(* IEC 61131-3 sources: ironplc/compiler/resources/test, 62 files *)

(* ---- first_steps_data_type_decl.st ---- *)
TYPE
  LOGLEVEL : (CRITICAL, WARNING, INFO, DEBUG) := INFO;
END_TYPE

(* ---- sized_string_contexts.st ---- *)
FUNCTION FUNC_WITH_VAR_STRING : INT
VAR_INPUT
    x : INT;
END_VAR
VAR
    buf : STRING[10];
    wbuf : WSTRING[20];
END_VAR
FUNC_WITH_VAR_STRING := 0;
END_FUNCTION

FUNCTION FUNC_WITH_VAR_CONSTANT_STRING : INT
VAR CONSTANT
    FILL : STRING[1] := '0';
    WFILL : WSTRING[1] := "0";
END_VAR
FUNC_WITH_VAR_CONSTANT_STRING := 0;
END_FUNCTION

FUNCTION FUNC_WITH_VAR_IN_OUT_STRING : INT
VAR_IN_OUT
    buf : STRING[255];
    wbuf : WSTRING[255];
END_VAR
FUNC_WITH_VAR_IN_OUT_STRING := 0;
END_FUNCTION

TYPE STRUCT_WITH_STRING :
STRUCT
    name : STRING[10];
    wname : WSTRING[20];
END_STRUCT;
END_TYPE

(* ---- strings.st ---- *)
TYPE
   TEXT_EXTENDED : STRING [1] := '�';
END_TYPE

(* ---- type_decl.st ---- *)
TYPE
   VALUES_ENUM : (VAL1, VAL2, VAL3);
   VALUES_ENUM_WITH_DEFAULT : (VAL1, VAL2, VAL3) := VAL2;
   LIMIT_RANGE : UINT (0..3);
   LIMIT_RANGE_DEFAULT : UINT (0..3) := 1;
   LIMIT_RANGE_NEGATIVE : INT(-10..10);
   ARR_RANGE : ARRAY[1..8] OF INT;
   ARR_RANGE_2D : ARRAY[1..8,1..4] OF INT;
   ARR_RANGE_ENUM : ARRAY[2..4] OF CUSTOM;
   TEXT_EMPTY : STRING [1];
   TEXT_DEFAULT : STRING [5] := 'value';
   WTEXT_EMPTY : WSTRING [1];
   WTEXT_DEFAULT : WSTRING [5] := 'value';
   CUSTOM_STRUCT : STRUCT
      NAME: BOOL;
   END_STRUCT;
   CUSTOM_STRUCT_WITH_ENUM : STRUCT
      NAME: VAL_TYPE := INIT_VAL;
      ARR_RANGE_ENUM : ARRAY[2..4] OF CUSTOM;
      LIMIT_RANGE : UINT (0..3);
      LIMIT_RANGE_DEFAULT : UINT (0..3) := 1;
   END_STRUCT;
   STR_WITH_SIZE : STRING[5];
   STR_WITH_SIZE_COMPATIBILITY : STRING[5];
END_TYPE

(* ---- array.st ---- *)
FUNCTION fun:BOOL

VAR_INPUT
    var1: INT;
    pt: ARRAY[1..8] OF INT;
END_VAR

var1 := var1 + pt[i];

END_FUNCTION

(* ---- array_in_function_var.st ---- *)
FUNCTION MY_FUNC : BOOL

VAR_INPUT
    x : INT;
END_VAR

VAR
    stack : ARRAY[1..32] OF UINT;
END_VAR

stack[1] := INT_TO_UINT(x);
MY_FUNC := TRUE;

END_FUNCTION

(* ---- array_of_string.st ---- *)
FUNCTION fun:BOOL

VAR_INPUT
    names: ARRAY[1..3] OF STRING[10];
END_VAR

fun := TRUE;

END_FUNCTION

(* ---- c_style_block_comment.st ---- *)
FUNCTION MY_FUNC : INT
VAR_INPUT
    x : INT;
END_VAR
    /* This is a C-style block comment */
    MY_FUNC := x;
END_FUNCTION

(* ---- empty_var_block.st ---- *)
FUNCTION myFunc : INT
VAR_INPUT
    x : INT;
END_VAR
VAR
END_VAR
    myFunc := x;
END_FUNCTION

(* ---- expressions.st ---- *)
FUNCTION fun:BOOL

VAR_INPUT
    var1: BYTE;
END_VAR

IF var1 < BYTE#32 THEN
	var1 := 1;
END_IF;

var1 := NOT (var3 OR var3);

var1 := FUNC_NAME(var1,'  ');

var1 := - 1 + 2 * 3 - 4 / 6 MOD 7 ** 8;

var1 := 1 >= 2 <= 3 <> 4 XOR 5;

IF var1 > t#1s THEN
    var1 := 1;
END_IF;

END_FUNCTION

(* ---- first_steps_func_avg_val.st ---- *)
FUNCTION AverageVal : REAL
    VAR_INPUT
    Cnt1 : INT;
    Cnt2 : INT;
    Cnt3 : INT;
    Cnt4 : INT;
    Cnt5 : INT;
  END_VAR
    VAR
    InputsNumber : REAL := 5.1;
  END_VAR
    AverageVal := INT_TO_REAL(Cnt1+Cnt2+Cnt3+Cnt4+Cnt5)/InputsNumber;
    END_FUNCTION

(* ---- inout_var_decl.st ---- *)
FUNCTION FUNC:UINT
    VAR_IN_OUT
        E : REAL;
        RNG : INT (1..2);
        ARR : ARRAY [0..3] OF INT;
    END_VAR

    array_avg := array_avg + arr[idx][idx];

END_FUNCTION

(* ---- input_var_decl.st ---- *)
FUNCTION FUNC:UINT
    VAR_INPUT
        E : REAL;
        PI, G : BOOL R_EDGE;
    END_VAR

    array_avg := array_avg + arr[idx][idx];

END_FUNCTION

(* ---- nested.st ---- *)
FUNCTION fun:BOOL

VAR_INPUT
    var1: BYTE;
END_VAR

array_avg := array_avg + arr[idx][idx];

END_FUNCTION

(* ---- bit_access.st ---- *)
FUNCTION_BLOCK MyBlock
  VAR
    myWord : WORD;
    myBool : BOOL;
  END_VAR

  myBool := myWord.0;
  myBool := myWord.15;
END_FUNCTION_BLOCK

(* ---- comment.st ---- *)
(* COMMENT *)
FUNCTION_BLOCK BLOCK
    (* MULTI-LINE
       COMMENT *)
    VAR_INT := 10;
END_FUNCTION_BLOCK

(* ---- conditional.st ---- *)
FUNCTION_BLOCK BLOCK

    IF NOT VAR1 AND VAR1 THEN
        VAR1 := 1;
    ELSIF NOT VAR1 AND VAR1 THEN
        VAR1 := 1;
    END_IF;

END_FUNCTION_BLOCK

(* ---- edge_input_decl.st ---- *)
FUNCTION_BLOCK Counter
    VAR_INPUT
        up : BOOL R_EDGE;
        down, reset : BOOL F_EDGE;
        amount : INT;
    END_VAR
    VAR_OUTPUT
        n : INT;
    END_VAR

    n := n + amount;

END_FUNCTION_BLOCK

PROGRAM main
    VAR_INPUT RETAIN
        go : BOOL R_EDGE;
    END_VAR
    VAR
        c : Counter;
    END_VAR

    c(up := go);

END_PROGRAM

(* ---- first_steps.st ---- *)
TYPE
  LOGLEVEL : (CRITICAL, WARNING, INFO, DEBUG) := INFO;
END_TYPE

FUNCTION_BLOCK LOGGER
  VAR_INPUT
    TRIG : BOOL;
    MSG : STRING;
    LEVEL : LOGLEVEL := INFO;
  END_VAR
  VAR
    TRIG0 : BOOL;
  END_VAR

  IF TRIG AND NOT TRIG0 THEN

  END_IF;
  TRIG0:=TRIG;
END_FUNCTION_BLOCK

FUNCTION_BLOCK CounterSFC
  VAR_INPUT
    Reset : BOOL;
  END_VAR
  VAR_OUTPUT
    OUT : INT;
  END_VAR
  VAR
    Cnt : INT;
  END_VAR
  VAR_EXTERNAL CONSTANT
    ResetCounterValue : INT;
  END_VAR

  INITIAL_STEP Start:
  END_STEP

  TRANSITION FROM Start TO ResetCounter
    := Reset;
  END_TRANSITION

  STEP ResetCounter:
    RESETCOUNTER_INLINE1(N);
    RESETCOUNTER_INLINE2(N);
  END_STEP

  ACTION RESETCOUNTER_INLINE1:
    Cnt := ResetCounterValue;
  END_ACTION

  ACTION RESETCOUNTER_INLINE2:
    OUT := Cnt;
  END_ACTION

  TRANSITION FROM ResetCounter TO Start
    := NOT Reset;
  END_TRANSITION

  TRANSITION FROM Start TO Count
    := NOT Reset;
  END_TRANSITION

  STEP Count:
    COUNT_INLINE3(N);
    COUNT_INLINE4(N);
  END_STEP

  ACTION COUNT_INLINE3:
    Cnt := Cnt + 1;
  END_ACTION

  ACTION COUNT_INLINE4:
    OUT := Cnt;
  END_ACTION

  TRANSITION FROM Count TO Start
    := Reset;
  END_TRANSITION

END_FUNCTION_BLOCK

FUNCTION_BLOCK CounterFBD
  VAR_INPUT
    Reset : BOOL;
  END_VAR
  VAR_OUTPUT
    OUT : INT;
  END_VAR
  VAR
    Cnt : INT;
  END_VAR
  VAR_EXTERNAL CONSTANT
    ResetCounterValue : INT;
  END_VAR
  VAR
    _TMP_ADD4_OUT : INT;
    _TMP_SEL7_OUT : INT;
  END_VAR

  Cnt := _TMP_SEL7_OUT;
  OUT := Cnt;
END_FUNCTION_BLOCK

FUNCTION AverageVal : REAL
  VAR_INPUT
    Cnt1 : INT;
    Cnt2 : INT;
    Cnt3 : INT;
    Cnt4 : INT;
    Cnt5 : INT;
  END_VAR
  VAR
    InputsNumber : REAL := 5.0;
  END_VAR

  AverageVal := INT_TO_REAL(Cnt1+Cnt2+Cnt3+Cnt4+Cnt5)/InputsNumber;
END_FUNCTION

FUNCTION_BLOCK CounterST
  VAR_INPUT
    Reset : BOOL;
  END_VAR
  VAR
    Cnt : INT;
  END_VAR
  VAR_OUTPUT
    OUT : INT;
  END_VAR
  VAR_EXTERNAL CONSTANT
    ResetCounterValue : INT;
  END_VAR

  IF Reset THEN
    Cnt := ResetCounterValue;
  ELSE
    Cnt := Cnt + 1;
  END_IF;

  Out := Cnt;
END_FUNCTION_BLOCK

FUNCTION_BLOCK CounterLD
  VAR_INPUT
    Reset : BOOL;
  END_VAR
  VAR_OUTPUT
    Out : INT;
  END_VAR
  VAR
    Cnt : INT;
  END_VAR
  VAR_EXTERNAL CONSTANT
    ResetCounterValue : INT;
  END_VAR
  VAR
    _TMP_ADD4_OUT : INT;
    _TMP_SEL7_OUT : INT;
  END_VAR

  Cnt := _TMP_SEL7_OUT;
  Out := Cnt;
END_FUNCTION_BLOCK

CONFIGURATION config
  VAR_GLOBAL CONSTANT
    ResetCounterValue : INT := 17;
  END_VAR

  RESOURCE resource1 ON PLC
    TASK plc_task(INTERVAL := T#100ms,PRIORITY := 1);
    PROGRAM plc_task_instance WITH plc_task : plc_prg;
  END_RESOURCE
END_CONFIGURATION

(* ---- first_steps_function_block_counter_fbd.st ---- *)
FUNCTION_BLOCK CounterFBD
  VAR_INPUT
    Reset : BOOL;
  END_VAR
  VAR_OUTPUT
    OUT : INT;
  END_VAR
  VAR
    Cnt : INT;
  END_VAR
  VAR_EXTERNAL CONSTANT
    ResetCounterValue : INT;
  END_VAR
  VAR
    _TMP_ADD4_OUT : INT;
    _TMP_SEL7_OUT : INT;
  END_VAR

  Cnt := _TMP_SEL7_OUT;
  OUT := Cnt;
END_FUNCTION_BLOCK

(* ---- first_steps_function_block_counter_ld.st ---- *)
FUNCTION_BLOCK CounterLD
  VAR_INPUT
    Reset : BOOL;
  END_VAR
  VAR_OUTPUT
    Out : INT;
  END_VAR
  VAR
    Cnt : INT;
  END_VAR
  VAR_EXTERNAL CONSTANT
    ResetCounterValue : INT;
  END_VAR
  VAR
    _TMP_ADD4_OUT : INT;
    _TMP_SEL7_OUT : INT;
  END_VAR

  _TMP_ADD4_OUT := ADD(1, Cnt);
  _TMP_SEL7_OUT := SEL(Reset, _TMP_ADD4_OUT, ResetCounterValue);
  Cnt := _TMP_SEL7_OUT;
  Out := Cnt;
END_FUNCTION_BLOCK

(* ---- first_steps_function_block_counter_sfc.st ---- *)
FUNCTION_BLOCK CounterSFC
  VAR_INPUT
    Reset : BOOL;
  END_VAR
  VAR_OUTPUT
    OUT : INT;
  END_VAR
  VAR
    Cnt : INT;
  END_VAR
  VAR_EXTERNAL CONSTANT
    ResetCounterValue : INT;
  END_VAR

  INITIAL_STEP Start:
  END_STEP

  TRANSITION FROM Start TO ResetCounter
    := Reset;
  END_TRANSITION

  STEP ResetCounter:
    RESETCOUNTER_INLINE1(N);
    RESETCOUNTER_INLINE2(N);
  END_STEP

  ACTION RESETCOUNTER_INLINE1:
    Cnt := ResetCounterValue;
  END_ACTION

  ACTION RESETCOUNTER_INLINE2:
    OUT := Cnt;
  END_ACTION

  TRANSITION FROM ResetCounter TO Start
    := NOT Reset;
  END_TRANSITION

  TRANSITION FROM Start TO Count
    := NOT Reset;
  END_TRANSITION

  STEP Count:
    COUNT_INLINE3(N);
    COUNT_INLINE4(N);
  END_STEP

  ACTION COUNT_INLINE3:
    Cnt := Cnt + 1;
  END_ACTION

  ACTION COUNT_INLINE4:
    OUT := Cnt;
  END_ACTION

  TRANSITION FROM Count TO Start
    := Reset;
  END_TRANSITION

END_FUNCTION_BLOCK

(* ---- first_steps_function_block_logger.st ---- *)
FUNCTION_BLOCK LOGGER
  VAR_INPUT
    TRIG : BOOL;
    MSG : STRING;
    LEVEL : LOGLEVEL := INFO;
  END_VAR
  VAR
    TRIG0 : BOOL;
  END_VAR

  IF TRIG AND NOT TRIG0 THEN

  END_IF;
  TRIG0:=TRIG;
END_FUNCTION_BLOCK

(* ---- first_steps_semantic_error.st ---- *)
TYPE
  LOGLEVEL : (CRITICAL, WARNING, INFO, DEBUG) := INFO;
END_TYPE

FUNCTION_BLOCK LOGGER
  VAR_INPUT
    TRIG : BOOL;
    MSG : STRING;
    LEVEL : LOGLEVEL := BLAH;
  END_VAR
  VAR
    TRIG0 : BOOL;
  END_VAR

  IF TRIG AND NOT TRIG0 THEN

  END_IF;
  TRIG0:=TRIG;
END_FUNCTION_BLOCK

FUNCTION_BLOCK CounterSFC
  VAR_INPUT
    Reset : BOOL;
  END_VAR
  VAR_OUTPUT
    OUT : INT;
  END_VAR
  VAR
    Cnt : INT;
  END_VAR
  VAR_EXTERNAL CONSTANT
    ResetCounterValue : INT;
  END_VAR

  INITIAL_STEP Start:
  END_STEP

  TRANSITION FROM Start TO ResetCounter
    := Reset;
  END_TRANSITION

  STEP ResetCounter:
    RESETCOUNTER_INLINE1(N);
    RESETCOUNTER_INLINE2(N);
  END_STEP

  ACTION RESETCOUNTER_INLINE1:
    Cnt := ResetCounterValue;
  END_ACTION

  ACTION RESETCOUNTER_INLINE2:
    OUT := Cnt;
  END_ACTION

  TRANSITION FROM ResetCounter TO Start
    := NOT Reset;
  END_TRANSITION

  TRANSITION FROM Start TO Count
    := NOT Reset;
  END_TRANSITION

  STEP Count:
    COUNT_INLINE3(N);
    COUNT_INLINE4(N);
  END_STEP

  ACTION COUNT_INLINE3:
    Cnt := Cnt + 1;
  END_ACTION

  ACTION COUNT_INLINE4:
    OUT := Cnt;
  END_ACTION

  TRANSITION FROM Count TO Start
    := Reset;
  END_TRANSITION

END_FUNCTION_BLOCK

FUNCTION_BLOCK CounterFBD
  VAR_INPUT
    Reset : BOOL;
  END_VAR
  VAR_OUTPUT
    OUT : INT;
  END_VAR
  VAR
    Cnt : INT;
  END_VAR
  VAR_EXTERNAL CONSTANT
    ResetCounterValue : INT;
  END_VAR
  VAR
    _TMP_ADD4_OUT : INT;
    _TMP_SEL7_OUT : INT;
  END_VAR

  Cnt := _TMP_SEL7_OUT;
  OUT := Cnt;
END_FUNCTION_BLOCK

FUNCTION AverageVal : REAL
  VAR_INPUT
    Cnt1 : INT;
    Cnt2 : INT;
    Cnt3 : INT;
    Cnt4 : INT;
    Cnt5 : INT;
  END_VAR
  VAR
    InputsNumber : REAL := 5.0;
  END_VAR

  AverageVal := INT_TO_REAL(Cnt1+Cnt2+Cnt3+Cnt4+Cnt5)/InputsNumber;
END_FUNCTION

FUNCTION_BLOCK CounterST
  VAR_INPUT
    Reset : BOOL;
  END_VAR
  VAR
    Cnt : INT;
  END_VAR
  VAR_OUTPUT
    OUT : INT;
  END_VAR
  VAR_EXTERNAL CONSTANT
    ResetCounterValue : INT;
  END_VAR

  IF Reset THEN
    Cnt := ResetCounterValue;
  ELSE
    Cnt := Cnt + 1;
  END_IF;

  Out := Cnt;
END_FUNCTION_BLOCK

FUNCTION_BLOCK CounterLD
  VAR_INPUT
    Reset : BOOL;
  END_VAR
  VAR_OUTPUT
    Out : INT;
  END_VAR
  VAR
    Cnt : INT;
  END_VAR
  VAR_EXTERNAL CONSTANT
    ResetCounterValue : INT;
  END_VAR
  VAR
    _TMP_ADD4_OUT : INT;
    _TMP_SEL7_OUT : INT;
  END_VAR

  Cnt := _TMP_SEL7_OUT;
  Out := Cnt;
END_FUNCTION_BLOCK

CONFIGURATION config
  VAR_GLOBAL CONSTANT
    ResetCounterValue : INT := 17;
  END_VAR

  RESOURCE resource1 ON PLC
    TASK plc_task(INTERVAL := T#100ms,PRIORITY := 1);
    PROGRAM plc_task_instance WITH plc_task : plc_prg;
  END_RESOURCE
END_CONFIGURATION

(* ---- first_steps_syntax_error.st ---- *)
TYPE
  LOGLEVEL : (CRITICAL, WARNING, INFO, DEBUG) := INFO;
END_TYPE

FUNCTION_BLOCK LOGGER
  VAR_INPUT
    TRIG : BOOL;
    MSG : STRING;
    LEVEL : LOGLEVEL := INFO;
  END_VAR
  VAR
    TRIG0 : BOOL;
  END_VAR

  IF TRIG AND NOT TRIG0 THEN

  END_IF;
  TRIG0:=TRIG;
END_FUNCTION_BLOCK

FUNCTION_BLOCK CounterSFC
  VAR_INPUT
    Reset : BOOL;
  END_VAR
  VAR_OUTPUT
    OUT : INT;
  END_VAR
  VAR
    Cnt : INT;
  END_VAR
  VAR_EXTERNAL CONSTANT
    ResetCounterValue : INT;
  END_VAR

  INITIAL_STEP Start:
  END_STEP

  TRANSITION FROM Start TO ResetCounter
    := Reset;
  END_TRANSITION

  STEP ResetCounter:
    RESETCOUNTER_INLINE1(N);
    RESETCOUNTER_INLINE2(N);
  END_STEP

  ACTION RESETCOUNTER_INLINE1:
    Cnt := ResetCounterValue;
  END_ACTION

  ACTION RESETCOUNTER_INLINE2:
    OUT := Cnt;
  END_ACTION

  TRANSITION FROM ResetCounter TO Start
    := NOT Reset;
  END_TRANSITION

  TRANSITION FROM Start TO Count
    := NOT Reset;
  END_TRANSITION

  STEP Count:
    COUNT_INLINE3(N);
    COUNT_INLINE4(N);
  END_STEP

  ACTION COUNT_INLINE3:
    Cnt := Cnt + 1;
  END_ACTION

  ACTION COUNT_INLINE4:
    OUT := Cnt;
  END_ACTION

  TRANSITION FROM Count TO Start
    := Reset;
  END_TRANSITION

END_FUNCTION_BLOCK

FUNCTION_BLOCK CounterFBD
  VAR_INPUT
    Reset : BOOL;
  END_VAR
  VAR_OUTPUT
    OUT : INT;
  END_VAR
  VAR
    Cnt : INT;
  END_VAR
  VAR_EXTERNAL CONSTANT
    ResetCounterValue : INT;
  END_VAR
  VAR
    _TMP_ADD4_OUT : INT;
    _TMP_SEL7_OUT : INT;
  END_VAR

  Cnt := _TMP_SEL7_OUT;
  OUT := Cnt;
END_FUNCTION_BLOCK

FUNCTION AverageVal : REAL
  VAR_INPUT
    Cnt1 : INT;
    Cnt2 : INT;
    Cnt3 : INT;
    Cnt4 : INT;
    Cnt5 : INT;
  END_VAR
  VAR
    InputsNumber : REAL := 5.0;
  END_VAR

  AverageVal := INT_TO_REAL(Cnt1+Cnt2+Cnt3+Cnt4+Cnt5)/InputsNumber;
END_FUNCTION

FUNCTION_BLOCK CounterST
  VAR_INPUT
    Reset : BOOL;
  END_VAR
  VAR
    Cnt : INT;
  END_VAR
  VAR_OUTPUT
    OUT : INT;
  END_VAR
  VAR_EXTERNAL CONSTANT
    ResetCounterValue : INT;
  END_VAR

  IF Reset THEN
    Cnt := ResetCounterValue;
  ELSE
    Cnt := Cnt + 1;
  END_IF;

  Out := Cnt;
END_FUNCTION_BLOCK

FUNCTION_BLOCK CounterLD
  VAR_INPUT
    Reset : BOOL
  END_VAR
  VAR_OUTPUT
    Out : INT;
  END_VAR
  VAR
    Cnt : INT;
  END_VAR
  VAR_EXTERNAL CONSTANT
    ResetCounterValue : INT;
  END_VAR
  VAR
    _TMP_ADD4_OUT : INT;
    _TMP_SEL7_OUT : INT;
  END_VAR

  Cnt := _TMP_SEL7_OUT;
  Out := Cnt;
END_FUNCTION_BLOCK

CONFIGURATION config
  VAR_GLOBAL CONSTANT
    ResetCounterValue : INT := 17;
  END_VAR

  RESOURCE resource1 ON PLC
    TASK plc_task(INTERVAL := T#100ms,PRIORITY := 1);
    PROGRAM plc_task_instance WITH plc_task : plc_prg;
  END_RESOURCE
END_CONFIGURATION

(* ---- if.st ---- *)
FUNCTION_BLOCK Error
    IF TRUE THEN
        Error := TRUE;
    END_IF
    IF TRUE THEN
        Error := TRUE;
    END_IF
END_FUNCTION_BLOCK

(* ---- literal.st ---- *)
FUNCTION_BLOCK BLOCK
    VAR
        REAL_WITH_TYPE: REAL := LREAL#11.0;
        BOOL_WITH_TYPE_TRUE: BOOL := BOOL#TRUE;
        TOD_WITH_VALUE_INTEGRAL: TIME_OF_DAY := TIME_OF_DAY#14:30:20;
        DATE_WITH_VALUE: DATE := DATE#2024-01-20;
        DATE_AND_TIME_WITH_VALUE: DATE_AND_TIME := DATE_AND_TIME#2024-01-20-15:30:22;
    END_VAR
    REAL_WITH_TYPE := 10;
END_FUNCTION_BLOCK

(* ---- oop.st ---- *)
INTERFACE I_Loggable
END_INTERFACE

INTERFACE I_Nameable
END_INTERFACE

INTERFACE I_Drivable EXTENDS I_Loggable
END_INTERFACE

FUNCTION_BLOCK ABSTRACT FB_BaseMotor IMPLEMENTS I_Drivable, I_Nameable
VAR
    bRunning : BOOL;
END_VAR
METHOD Start
    bRunning := TRUE;
END_METHOD
METHOD Stop
    bRunning := FALSE;
END_METHOD
END_FUNCTION_BLOCK

FUNCTION_BLOCK FB_ServoMotor EXTENDS FB_BaseMotor IMPLEMENTS I_Drivable
VAR
    rSpeed : REAL;
    aHistory : ARRAY[0..3] OF REAL;
END_VAR
METHOD SetSpeed : BOOL
VAR_INPUT
    rNewSpeed : REAL;
END_VAR
    SUPER^.Start();
    rSpeed := rNewSpeed;
    THIS^.aHistory[0] := rNewSpeed;
    SetSpeed := TRUE;
END_METHOD
METHOD LogState
    IF SUPER^.bRunning THEN
        aHistory[1] := rSpeed;
    END_IF;
END_METHOD
METHOD Reset
    THIS^.rSpeed := 0.0;
    THIS^.LogState();
    SUPER^.Stop();
END_METHOD
END_FUNCTION_BLOCK

PROGRAM main
VAR
    m : FB_ServoMotor;
END_VAR
m.SetSpeed(1.5);
m.SetSpeed(rNewSpeed := 2.0);
m.Reset();
END_PROGRAM

(* ---- partial_access_bit.st ---- *)
FUNCTION_BLOCK MyBlock
  VAR
    myWord : WORD;
    myBool : BOOL;
  END_VAR

  myBool := myWord.%X0;
  myBool := myWord.%X15;
END_FUNCTION_BLOCK

(* ---- sfc.st ---- *)
FUNCTION_BLOCK sfc
  VAR_INPUT
    IN : BOOL;
  END_VAR
  VAR_OUTPUT
    OUT : INT;
  END_VAR
  VAR
    COUNT : INT;
  END_VAR

  INITIAL_STEP Start:
    RESET(N);
  END_STEP

  TRANSITION FROM Start TO MidStep
    := FALSE;
  END_TRANSITION

  STEP MidStep:
    RESET(N);
  END_STEP

  ACTION RESET:
    COUNT := 0;
  END_ACTION

END_FUNCTION_BLOCK

(* ---- textual.st ---- *)
FUNCTION_BLOCK BLOCK
    NUM_INT := 10;
    NUM_FLOAT := 10.0;

    IF NUM1 < NUM2 THEN
        NUM1 := 1;
    ELSIF NUM2 = NUM3 THEN
        NUM1 := 2;
    ELSE
        NUM1 := 3;
    END_IF;

    CASE EXPR_WITH_ELSE OF
    VAL1: (* empty *);
    VAL2: NUM1 := 1;
    ELSE NUM2 := 2;
    END_CASE;

    CASE EXPR_NO_ELSE OF
    VAL1: (* empty *);
    VAL2: NUM1 := 1;
    END_CASE;

    FOR VAL1 := 1 TO 10 BY 1 DO
       VAL2 := VAL1;
    END_FOR;

    WHILE VAL1 = 1 DO
        VAL2 := VAL1;
    END_WHILE;

    REPEAT
        VAL2 := VAL1;
    UNTIL VAL2 = 2
    END_REPEAT;

END_FUNCTION_BLOCK

(* ---- try_catch.st ---- *)
(* CODESYS exception handling: __TRY/__CATCH/__FINALLY/__ENDTRY, __THROW. *)

PROGRAM main
VAR
    e : INT;
    x : INT;
END_VAR
    __TRY
        x := 1;
        IF x > 0 THEN
            __THROW(7);
        END_IF;
        x := 2;
    __CATCH (e)
        x := e;
    __FINALLY
        x := x + 1;
    __ENDTRY;
END_PROGRAM

FUNCTION_BLOCK guarded
VAR
    n : INT;
END_VAR
    __TRY
        n := n + 1;
    __ENDTRY;
    __TRY
        n := n + 2;
    __FINALLY
        n := n + 3;
    __ENDTRY;
    __TRY
        n := n + 4;
    __CATCH ()
        n := 0;
    __ENDTRY;
    __TRY
        n := n + 5;
    __CATCH
        __THROW;
    __ENDTRY;
END_FUNCTION_BLOCK

(* ---- typed_string_literals.st ---- *)
FUNCTION_BLOCK typed_literals
VAR
    narrow : STRING[20];
    wide : WSTRING[20];
    code : STRING[20];
END_VAR
    narrow := UTF8#'a$41b';
    wide := __XSTRING#"a$0041b";
    code := UCHAR#'A';
END_FUNCTION_BLOCK

(* ---- var_sections.st ---- *)
(* CODESYS/TwinCAT additional variable sections: VAR_STAT (static),
   VAR_INST (method instance) and VAR_GENERIC (function block generic
   constants). Parsed with the CODESYS dialect. *)

FUNCTION CountUp : DINT
VAR_STAT
    calls : DINT;
END_VAR
    calls := calls + 1;
    CountUp := calls;
END_FUNCTION

FUNCTION_BLOCK FB_Scale
VAR_GENERIC CONSTANT
    maxValue : INT := 100;
END_VAR
VAR
    value : INT;
END_VAR
    value := maxValue;
METHOD Clamp : INT
VAR_INST
    clamped : INT;
END_VAR
    IF value > maxValue THEN
        clamped := maxValue;
    ELSE
        clamped := value;
    END_IF;
    Clamp := clamped;
END_METHOD
END_FUNCTION_BLOCK

PROGRAM main
VAR_STAT
    scans : DINT;
END_VAR
VAR
    scale : FB_Scale;
    result : INT;
END_VAR
    scans := scans + 1;
    result := scale.Clamp();
END_PROGRAM

(* ---- var_temp.st ---- *)
FUNCTION my_func : DINT
  VAR_INPUT
    a : DINT;
  END_VAR
  VAR_TEMP
    temp : DINT;
  END_VAR
  temp := a * 2;
  my_func := temp;
END_FUNCTION

FUNCTION_BLOCK my_fb
  VAR_TEMP
    t : INT;
  END_VAR
  t := 42;
END_FUNCTION_BLOCK

PROGRAM my_prog
  VAR_TEMP
    t : INT;
  END_VAR
  t := 7;
END_PROGRAM

(* ---- adr.st ---- *)
PROGRAM main
VAR
    counter : INT := 42;
    p : POINTER TO INT;
    value : INT;
END_VAR
    p := ADR(counter);
    value := p^;
    p^ := 99;
END_PROGRAM

(* ---- based_literals.st ---- *)
PROGRAM main
VAR
    x : DINT;
    b : BOOL;
    one : BIT;
END_VAR
    x := 10#123;
    b := BOOL#1;
    one := BIT#1;
END_PROGRAM

(* ---- bit_string_arithmetic.st ---- *)
(* Arithmetic on a bit-string operand: accepted only with
   --allow-bit-string-arithmetic or a dialect that enables it. *)
PROGRAM main
  VAR
    counter : BYTE;
  END_VAR
  counter := counter + 1;
END_PROGRAM

(* ---- case_selectors.st ---- *)
TYPE
    E_State : (Idle, Run, Stop);
END_TYPE

PROGRAM main
    VAR
        n : INT;
        s : E_State;
        x : INT;
    END_VAR

    CASE n OF
        1, 2: x := 1;
        3..5: x := 2;
        6, 8..9, 12: x := 3;
        ELSE x := 4;
    END_CASE;

    CASE s OF
        Idle, E_State#Run: x := 5;
        Stop: x := 6;
    END_CASE;
END_PROGRAM

(* ---- configuration.st ---- *)
CONFIGURATION config
  RESOURCE resource1 ON PLC
    TASK plc_task(INTERVAL := T#100ms,PRIORITY := 1);
    PROGRAM plc_task_instance WITH plc_task : plc_prg;
  END_RESOURCE

  VAR_CONFIG
    Some.Located.Item.Path AT %QB1: BYTE;
    Some.FunctionBlock.Item.Path : FB_TYPE_NAME := (ELEM := VAL);
  END_VAR
END_CONFIGURATION

PROGRAM main
    VAR
        Button AT %IX1: BOOL;
        Buzzer AT %QX1: BOOL;
    END_VAR

    Buzzer := NOT Button;

END_PROGRAM

(* ---- escaped_identifiers.st ---- *)
PROGRAM main
VAR
    `counter value` : INT;
    `CAFÉ` : INT;
END_VAR
    `counter value` := 1;
    `CAFÉ` := 2;
END_PROGRAM

(* ---- first_steps_configuration.st ---- *)
CONFIGURATION config
  VAR_GLOBAL CONSTANT
    ResetCounterValue : INT := 17;
  END_VAR

  RESOURCE resource1 ON PLC
    TASK plc_task(INTERVAL := T#100ms,PRIORITY := 1);
    PROGRAM plc_task_instance WITH plc_task : plc_prg;
  END_RESOURCE
END_CONFIGURATION

(* ---- first_steps_program.st ---- *)
PROGRAM plc_prg
  VAR_INPUT
    Reset : BOOL;
  END_VAR
  VAR_OUTPUT
    Cnt1 : INT;
    Cnt2 : INT;
    Cnt3 : INT;
    Cnt4 : INT;
    Cnt5 : INT;
  END_VAR
  VAR
    CounterST0 : CounterST;
    CounterFBD0 : CounterFBD;
    CounterSFC0 : CounterSFC;
    CounterIL0 : CounterIL;
    CounterLD0 : CounterLD;
    AVCnt : REAL;
    _TMP_AverageVal17_OUT : REAL;
  END_VAR

  CounterST0(Reset := Reset);
  Cnt1 := CounterST0.OUT;
  _TMP_AverageVal17_OUT := AverageVal(Cnt1, Cnt2, Cnt3, Cnt4, Cnt5);
  AVCnt := _TMP_AverageVal17_OUT;
  CounterFBD0(Reset := Reset);
  Cnt2 := CounterFBD0.OUT;
  CounterSFC0(Reset := Reset);
  Cnt3 := CounterSFC0.OUT;
  CounterIL0(Reset := Reset);
  Cnt4 := CounterIL0.OUT;
  CounterLD0(Reset := Reset);
  Cnt5 := CounterLD0.Out;
END_PROGRAM

(* ---- incomplete_array.st ---- *)
TYPE DataBuffer : ARRAY[*] OF INT; END_TYPE

PROGRAM main
VAR
    data : ARRAY[*] OF BYTE;
END_VAR
END_PROGRAM

(* ---- main.st ---- *)
   PROGRAM main
      VAR
         Button AT %IX1: BOOL;
         Buzzer AT %QX1: BOOL;
      END_VAR

      Buzzer := NOT Button;

   END_PROGRAM

   CONFIGURATION config
      RESOURCE res ON PLC
         TASK plc_task(INTERVAL := T#100ms, PRIORITY := 1);
         PROGRAM plc_task_instance WITH plc_task : main;
      END_RESOURCE
   END_CONFIGURATION

(* ---- namespace.st ---- *)
(* CODESYS/TwinCAT NAMESPACE grouping plus the __BEGIN_IMPLEMENTATION
   implementation marker. Parsed with --allow-namespace and
   --allow-begin-implementation (the CODESYS dialect enables both). *)

NAMESPACE Motor
TYPE
E_Direction : (Forward, Backward);
END_TYPE

FUNCTION Blocked : BOOL
VAR_INPUT
    dir : INT;
END_VAR
    Blocked := dir < 0;
END_FUNCTION

NAMESPACE Control
PROGRAM main
VAR
    moving : BOOL;
END_VAR
__BEGIN_IMPLEMENTATION
    moving := NOT Blocked(1);
END_PROGRAM
END_NAMESPACE
END_NAMESPACE

(* ---- oscat.st ---- *)
(*@PROPERTIES_EX@
TYPE: POU
LOCALE: 0
IEC_LANGUAGE: ST
PLC_TYPE: independent
PROC_TYPE: independent
GROUP:
*)
(*@KEY@:DESCRIPTION*)
version 1.0	1. jan. 2000
programmer 	garret
tested by	garret

some description
(*@KEY@:END_DESCRIPTION*)
TYPE
    CUSTOM_STRUCT : STRUCT
        NAME: BOOL;
    END_STRUCT;
END_TYPE

(* ---- params_of.st ---- *)
TYPE ScaledParams : PARAMS(2) OF REAL; END_TYPE

PROGRAM main
VAR
    args : PARAMS(3) OF INT;
    named : ScaledParams;
END_VAR
    args[0] := 1;
END_PROGRAM

(* ---- partial_access_multi.st ---- *)
PROGRAM main
  VAR
    d : DWORD;
    l : LWORD;
    rb : BYTE;
    rw : WORD;
    rd : DWORD;
  END_VAR
  rb := d.%B0;
  rw := d.%W1;
  rd := l.%D0;
  d.%B2 := BYTE#16#FF;
  l.%W3 := WORD#16#ABCD;
END_PROGRAM

(* ---- pipe_or.st ---- *)
PROGRAM main
VAR
    a : BOOL;
    b : BOOL;
    c : BOOL;
    or_result : BOOL;
    mixed : BOOL;
END_VAR
    or_result := a | b;
    mixed := a | b & c;
END_PROGRAM

(* ---- pointer_to.st ---- *)
TYPE IntPtr : POINTER TO INT; END_TYPE

PROGRAM main
VAR
    counter : INT := 42;
    p : POINTER TO INT;
    ptrs : ARRAY[0..2] OF POINTER TO INT;
    value : INT;
END_VAR
    p := REF(counter);
    value := p^;
    p^ := 99;
    p := NULL;
END_PROGRAM

(* ---- program.st ---- *)
PROGRAM main
    VAR
        Button AT %IX1: BOOL;
        Buzzer AT %QX1: BOOL;
    END_VAR
    VAR_ACCESS
        VarPath : VarName.Path : BOOL READ_ONLY;
    END_VAR

    Buzzer := NOT Button;

END_PROGRAM

(* ---- ref.st ---- *)
TYPE IntRef : REF_TO INT; END_TYPE

TYPE ArrRef : REF_TO ARRAY[0..3] OF DINT; END_TYPE

FUNCTION read_ref : INT
VAR_INPUT
    pt : REF_TO INT;
END_VAR
    read_ref := pt^;
END_FUNCTION

PROGRAM main
VAR
    counter : INT := 42;
    r : REF_TO INT := REF(counter);
    r_null : REF_TO INT := NULL;
    r_uninit : REF_TO INT;
    data : REF_TO ARRAY[0..3] OF INT;
    refs : ARRAY[0..2] OF REF_TO INT;
    value : INT;
END_VAR
    value := r^;
    r^ := 99;
    r := REF(counter);
    IF r <> NULL THEN
        value := r^;
    END_IF;
    value := read_ref(pt := REF(counter));
END_PROGRAM

(* ---- reference_to.st ---- *)
TYPE IntRef : REFERENCE TO INT; END_TYPE

PROGRAM main
VAR
    counter : INT := 42;
    r : REFERENCE TO INT;
    refs : ARRAY[0..2] OF REFERENCE TO INT;
    value : INT;
END_VAR
    r REF= counter;
    value := r^;
    r^ := 99;
    refs[0] REF= counter;
    value := refs[0]^;
END_PROGRAM

(* ---- sizeof.st ---- *)
PROGRAM main
VAR
  x : INT;
  y : DWORD;
  arr : ARRAY[1..10] OF INT;
  s : DINT;
END_VAR
  s := SIZEOF(x);
  s := SIZEOF(y);
  s := SIZEOF(arr);
END_PROGRAM

(* ---- special_operators.st ---- *)
PROGRAM main
VAR
    result : DINT;
    obj : INT;
END_VAR
    obj := __NEW(INT);
    obj := __NEW(INT, 4);
    result := __XADD(1, 2);
    result := __DELETE(obj);
    result := __TYPEOF(DINT);
    result := __ISVALIDREF(obj);
END_PROGRAM

(* ---- steel_thread.st ---- *)
PROGRAM main
  VAR
    x : INT;
    y : INT;
  END_VAR
  x := 10;
  y := x + 32;
END_PROGRAM

(* ---- time_function_decl.st ---- *)
FUNCTION TIME : TIME
TIME := T#0s;
END_FUNCTION

PROGRAM main
VAR
    t : TIME;
END_VAR
t := TIME();
END_PROGRAM

(* ---- time_literal_extensions.st ---- *)
PROGRAM main
VAR
    micro : TIME := T#1us;
    nano : TIME := T#500ns;
    long : LTIME := LT#1500us;
    fraction : TIME := T#1.5ms;
    day : DATE := LD#2024-01-20;
    clock : TIME_OF_DAY := TOD#10:00;
END_VAR
END_PROGRAM

(* ---- union.st ---- *)
(* CODESYS UNION type declaration (IEC 61131-3:2013).
   Parsed with --allow-union-type / --dialect codesys. *)
TYPE
U_Data :
UNION
    intVal : INT;
    realVal : REAL;
    flags : ARRAY[0..31] OF BOOL;
END_UNION;
U_Point :
UNION
    x : INT := 1;
    pair : ARRAY[0..1] OF INT;
END_UNION;
END_TYPE

PROGRAM main
VAR
    data : U_Data;
    x : INT;
END_VAR
    data.intVal := 1;
    x := data.intVal;
END_PROGRAM

(* ---- var_decl.st ---- *)
PROGRAM fb
    VAR CONSTANT
        E : REAL := 2.718 ;
    END_VAR

    VAR
        AT %IX1.1 : BOOL;
        AT %IX2.1 : BOOL :=1;
        AT %MW1 : INT := 2 ;
    END_VAR

    VAR RETAIN
       AT %QW1 : WORD := 16#FF00 ;
       AT %QB2 : WORD := 8#7700 ;
       AT %QB3 : WORD := 2#1010 ;
       C3 AT %MW1.2.3 : WORD;
    END_VAR

    VAR RETAIN
        C2 AT %Q* : BYTE ;
    END_VAR

    VAR
        XWORD, YWORD, ZWORD : INT;

        UNINIT: ARRAY [0..9] OF INT;
        INIT : ARRAY [1..12] OF SINT := [2,7,18];
        MULTI_DIM_ARRAY : ARRAY[1..2,3..4,5..6] OF SINT;
        PARENTHESIS_ARRAY : ARRAY[0..3] OF SINT := [3(2)];

        VAL_STR: STRING[2];
        VAL_STR_INIT: STRING := 'abc';
        VAL_STR_PREFIX: STRING := STRING#'ABC';
        VAL_STR_SIZED_INIT: STRING[3] := 'abc';
        VAL_WSTR: WSTRING[9];
        VAL_WSTR_INIT: WSTRING := "def";
        VAL_WSTR_PREFIX: WSTRING := WSTRING#"ABC";
        VAL_WSTR_SIZED_INIT: WSTRING[3] := "def";
    END_VAR

    VAR
        NAME : ONE_STRUCT_ELEMENT := (ELEM := VAL);
        NAME2 : TWO_STRUCT_ELEMENTS := (ELEM1 := VAL1, ELEM2 := VAL2);
        NAME3 : STRUCT_TWO_ELEMENTS := (ELEM1 := VAL1, ELEM2 := VAL2);
        (* TODO Nested structures *)
    END_VAR

    VAR
		X :	REAL2;
		Y :	REAL;
	END_VAR

END_PROGRAM

(* ---- wstring_ops.st ---- *)
PROGRAM main
    VAR
        a : WSTRING[10] := "foo";
        b : WSTRING[10] := "bar";
        c : WSTRING[20];
        s : STRING[20];
        n : DINT;
        eq : BOOL;
    END_VAR
    c := a;
    c := "baz";
    s := 'baz';
    c := CONCAT(a, b);
    n := LEN(a);
    eq := a = b;
END_PROGRAM
